FUNCTION F_JsonNumSigned : BOOL
VAR_INPUT
    sKey      : STRING(31);
    fValue    : LREAL;
    bValid    : BOOL;
    nDecimals : INT;  // 0..3
END_VAR
VAR_IN_OUT
    fbJson : FB_JsonSaxWriter;
END_VAR
VAR
    fTmp   : LREAL;
    fScale : LREAL;
    bOk    : BOOL;
END_VAR

fTmp := fValue;
bOk := FALSE;
IF bValid THEN
    IF IsFinite(F_LREAL(fTmp)) THEN
        bOk := ABS(fTmp) < 1.0E12;
    END_IF
END_IF

fbJson.AddKey(sKey);
IF bOk THEN
    CASE nDecimals OF
        1: fScale := 10.0;
        2: fScale := 100.0;
        3: fScale := 1000.0;
    ELSE
        fScale := 1.0;
    END_CASE
    fbJson.AddLreal(LINT_TO_LREAL(LREAL_TO_LINT(fTmp * fScale)) / fScale);
ELSE
    fbJson.AddNull();
END_IF
F_JsonNumSigned := bOk;

END_FUNCTION

(* stored: Version 1.1.0.1
   POU F_JsonNumSigned: Id {1ad9fd1f-ba22-435e-a844-92f625a25329}, SpecialFunc None *)
